(* Logix 5000 project; controller TFF vendor 1 type 14 code 107 rev 33.11; software revision 33.04; part 35 of 38 *)
(* tags used below, declared in another part *)
   Index : DINT;   // Index
   TIME : DINT[2];
   DigitalOutput : BOOL[256];   // Digital Output Array these bits are sent to output cards.
   FlowPath : FlowPath[64];   // Flow Path Array
   Options : Options;   // Options List
   PCV101_Control : PCV_Control;   // PCV101 Control UDT
   PCV201_Control : PCV_Control;   // PCV201 Control UDT
   PipeAnimation : PipeAnimation;   // HMI Pipe Animation Array
   PipeStatValueHMI : INT[224];   // Pipe Animation Value For HMI
   PTA001 : ALIAS FOR DigitalOutput[21];
   PTA101 : ALIAS FOR DigitalOutput[22];
   PTA201 : ALIAS FOR DigitalOutput[23];
   PTA401 : ALIAS FOR DigitalOutput[24];
   Rack_Murr_Node1_TFF20 : IO_Station;   // Status of Node 1 TFF20
   ThisSystem : SystemType;
   XV001 : ALIAS FOR Valve[0];
   XV002 : ALIAS FOR Valve[1];
   XV003 : ALIAS FOR Valve[2];
   XV004 : ALIAS FOR Valve[3];
   XV005 : ALIAS FOR Valve[4];
   XV006 : ALIAS FOR Valve[5];
   XV007 : ALIAS FOR Valve[6];
   XV101 : ALIAS FOR Valve[7];
   XV102 : ALIAS FOR Valve[8];
   XV201 : ALIAS FOR Valve[15];
   XV202 : ALIAS FOR Valve[16];
   XV401 : ALIAS FOR Valve[9];
   XV402 : ALIAS FOR Valve[10];
   XV403 : ALIAS FOR Valve[11];
   XV404 : ALIAS FOR Valve[12];
   XV405 : ALIAS FOR Valve[13];
   XV406 : ALIAS FOR Valve[14];
   XV701 : ALIAS FOR Valve[17];
   XV702 : ALIAS FOR Valve[18];
   XV703 : ALIAS FOR Valve[19];
   XV704 : ALIAS FOR Valve[20];
(* Process, continued *)

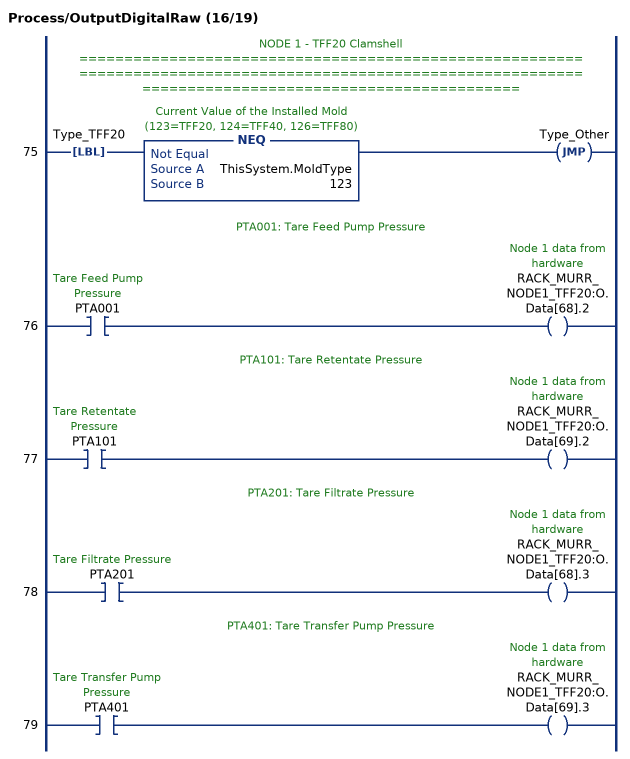
   // NODE 1 - TFF20 Clamshell
   // ==========================================================================================================================================================
   75: LBL(Type_TFF20)NEQ(ThisSystem.MoldType,123)JMP(Type_Other);
   // PTA001: Tare Feed Pump Pressure
   76: XIC(PTA001)OTE(RACK_MURR_NODE1_TFF20:O.Data[68].2);
   // PTA101: Tare Retentate Pressure
   77: XIC(PTA101)OTE(RACK_MURR_NODE1_TFF20:O.Data[69].2);
   // PTA201: Tare Filtrate Pressure
   78: XIC(PTA201)OTE(RACK_MURR_NODE1_TFF20:O.Data[68].3);
   // PTA401: Tare Transfer Pump Pressure
   79: XIC(PTA401)OTE(RACK_MURR_NODE1_TFF20:O.Data[69].3);
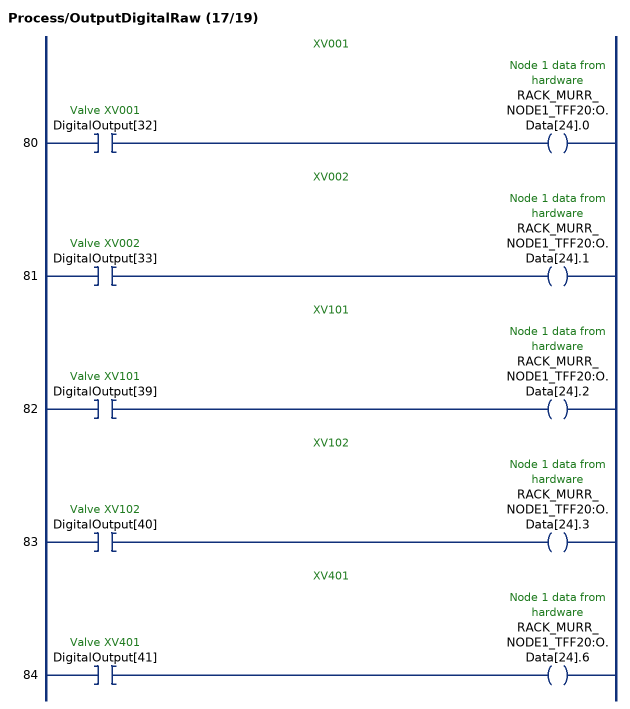
   // XV001
   80: XIC(DigitalOutput[32])OTE(RACK_MURR_NODE1_TFF20:O.Data[24].0);
   // XV002
   81: XIC(DigitalOutput[33])OTE(RACK_MURR_NODE1_TFF20:O.Data[24].1);
   // XV101
   82: XIC(DigitalOutput[39])OTE(RACK_MURR_NODE1_TFF20:O.Data[24].2);
   // XV102
   83: XIC(DigitalOutput[40])OTE(RACK_MURR_NODE1_TFF20:O.Data[24].3);
   // XV401
   84: XIC(DigitalOutput[41])OTE(RACK_MURR_NODE1_TFF20:O.Data[24].6);
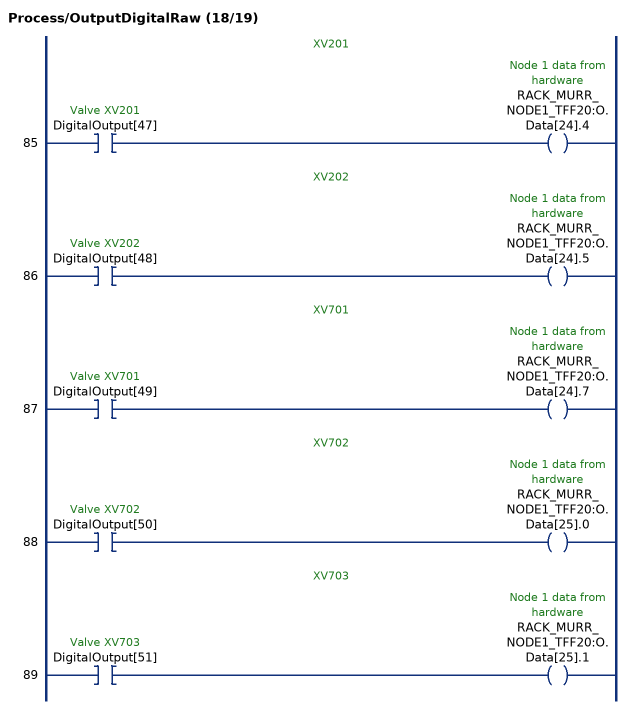
   // XV201
   85: XIC(DigitalOutput[47])OTE(RACK_MURR_NODE1_TFF20:O.Data[24].4);
   // XV202
   86: XIC(DigitalOutput[48])OTE(RACK_MURR_NODE1_TFF20:O.Data[24].5);
   // XV701
   87: XIC(DigitalOutput[49])OTE(RACK_MURR_NODE1_TFF20:O.Data[24].7);
   // XV702
   88: XIC(DigitalOutput[50])OTE(RACK_MURR_NODE1_TFF20:O.Data[25].0);
   // XV703
   89: XIC(DigitalOutput[51])OTE(RACK_MURR_NODE1_TFF20:O.Data[25].1);
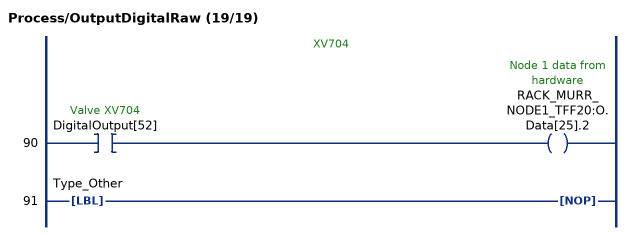
   // XV704
   90: XIC(DigitalOutput[52])OTE(RACK_MURR_NODE1_TFF20:O.Data[25].2);
   91: LBL(Type_Other)NOP();
END_ROUTINE

ROUTINE OutputProcessing   (* ladder *)
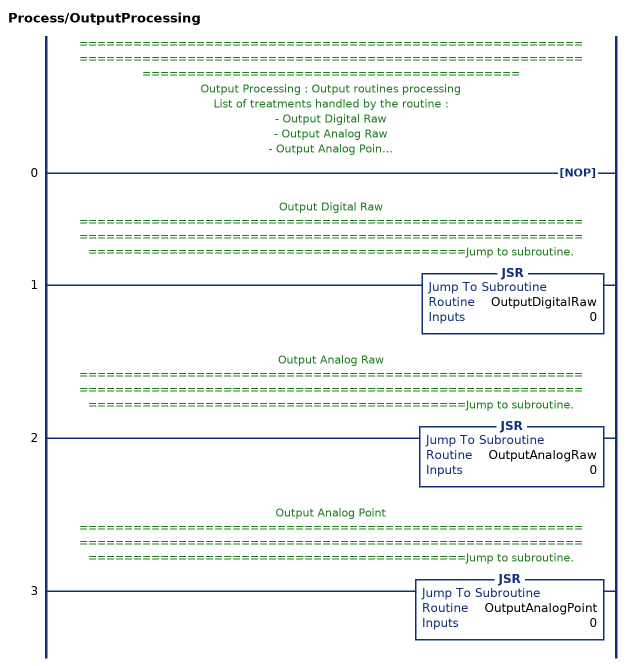
   // ==========================================================================================================================================================
   //                                                                                                                  Output Processing : Output routines processing
   //                                                     List of treatments handled by the routine :
   //                                                          - Output Digital Raw
   //                                                          - Output Analog Raw
   //                                                          - Output Analog Point
   //                                                     -----------------------------------------------------------------------------------------------------------------------------------------------------
   //                                                     History
   // 		2019-DEC-24 - Merck - Q. Spindler - Initial version for Candidate Release 1.00.00.00.a
   // ==========================================================================================================================================================
   0: NOP();
   // Output Digital Raw
   // ==========================================================================================================================================================Jump to subroutine.
   1: JSR(OutputDigitalRaw,0);
   // Output Analog Raw
   // ==========================================================================================================================================================Jump to subroutine.
   2: JSR(OutputAnalogRaw,0);
   // Output Analog Point
   // ==========================================================================================================================================================Jump to subroutine.
   3: JSR(OutputAnalogPoint,0);
END_ROUTINE

ROUTINE PipeAnimation   (* ladder *)
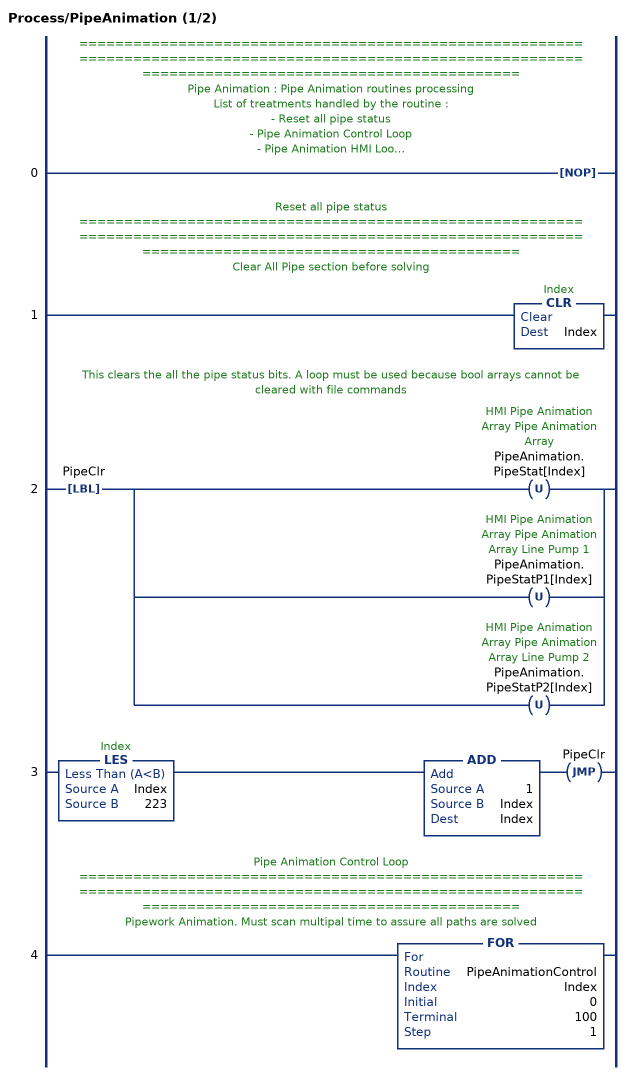
   // ==========================================================================================================================================================
   //                                                                                                               Pipe Animation : Pipe Animation routines processing
   //                                                     List of treatments handled by the routine :
   //                                                          - Reset all pipe status
   //                                                          - Pipe Animation Control Loop
   //                                                          - Pipe Animation HMI Loop
   //                                                     -----------------------------------------------------------------------------------------------------------------------------------------------------
   //                                                     History
   // 		2019-DEC-24 - Merck - Q. Spindler - Initial version for Candidate Release 1.00.00.00.a
   // ==========================================================================================================================================================
   0: NOP();
   // Reset all pipe status
   // ==========================================================================================================================================================
   // Clear All Pipe section before solving
   1: CLR(Index);
   // This clears the all the pipe status bits. A loop must be used because bool arrays cannot be cleared with file commands
   2: LBL(PipeClr)[OTU(PipeAnimation.PipeStat[Index]) ,OTU(PipeAnimation.PipeStatP1[Index]) ,OTU(PipeAnimation.PipeStatP2[Index]) ];
   3: LES(Index,223)ADD(1,Index,Index)JMP(PipeClr);
   // Pipe Animation Control Loop
   // ==========================================================================================================================================================
   // Pipework Animation. Must scan multipal time to assure all paths are solved
   4: FOR(PipeAnimationControl,Index,0,100,1);
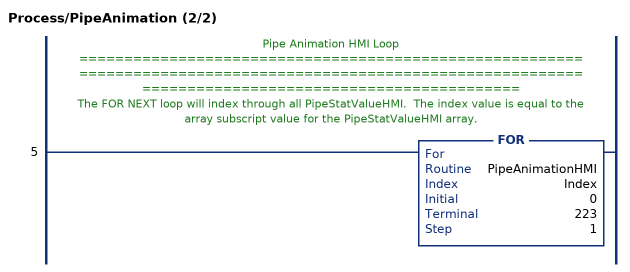
   // Pipe Animation HMI Loop
   // ==========================================================================================================================================================
   // The FOR NEXT loop will index through all PipeStatValueHMI.  The index value is equal to the array subscript value for the PipeStatValueHMI array.
   5: FOR(PipeAnimationHMI,Index,0,223,1);
END_ROUTINE

ROUTINE PipeAnimationControl   (* ladder *)
// Pipework Animation Routine
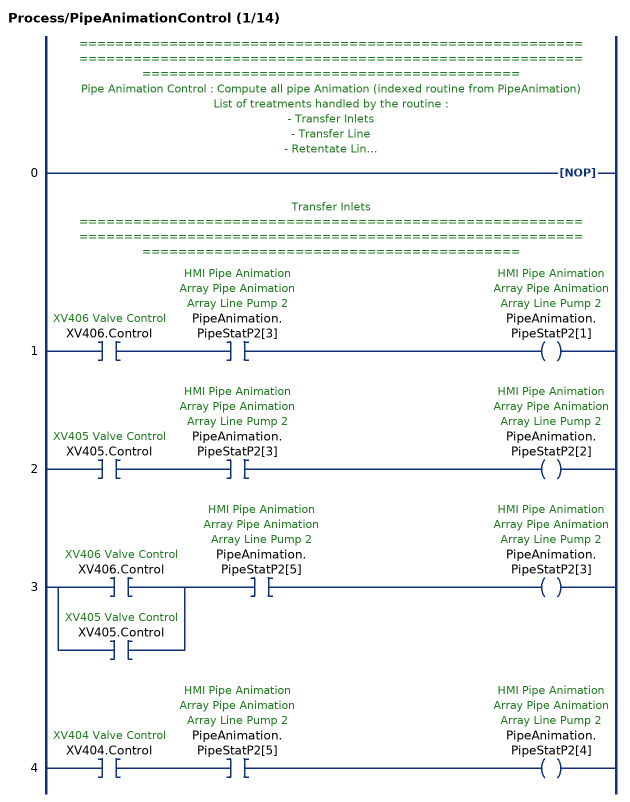
   // ==========================================================================================================================================================
   //                                                                                        Pipe Animation Control : Compute all pipe Animation (indexed routine from PipeAnimation)
   //                                                     List of treatments handled by the routine :
   //                                                          - Transfer Inlets
   //                                                          - Transfer Line
   //                                                          - Retentate Line
   //                                                           - Filtrate
   //                                                          - Feed Line
   //                                                           - Feed Inlets
   //                                                     -----------------------------------------------------------------------------------------------------------------------------------------------------
   //                                                     History
   // 		2019-DEC-24 - Merck - Q. Spindler - Initial version for Candidate Release 1.00.00.00.a
   // 		2020-JUN-19 - Merck - Q. Spindler - Modifications for Candidate Release 1.00.00.00.c
   //                                                                                             - Change State for Pipe ID 13, 14, 15, 16, 17, and 18 to prohibit Frontal filtration flowpath
   // ========================================================================================================================================================
   0: NOP();
   // Transfer Inlets
   // ==========================================================================================================================================================
   1: XIC(XV406.Control)XIC(PipeAnimation.PipeStatP2[3])OTE(PipeAnimation.PipeStatP2[1]);
   2: XIC(XV405.Control)XIC(PipeAnimation.PipeStatP2[3])OTE(PipeAnimation.PipeStatP2[2]);
   3: [XIC(XV406.Control) ,XIC(XV405.Control) ]XIC(PipeAnimation.PipeStatP2[5])OTE(PipeAnimation.PipeStatP2[3]);
   4: XIC(XV404.Control)XIC(PipeAnimation.PipeStatP2[5])OTE(PipeAnimation.PipeStatP2[4]);
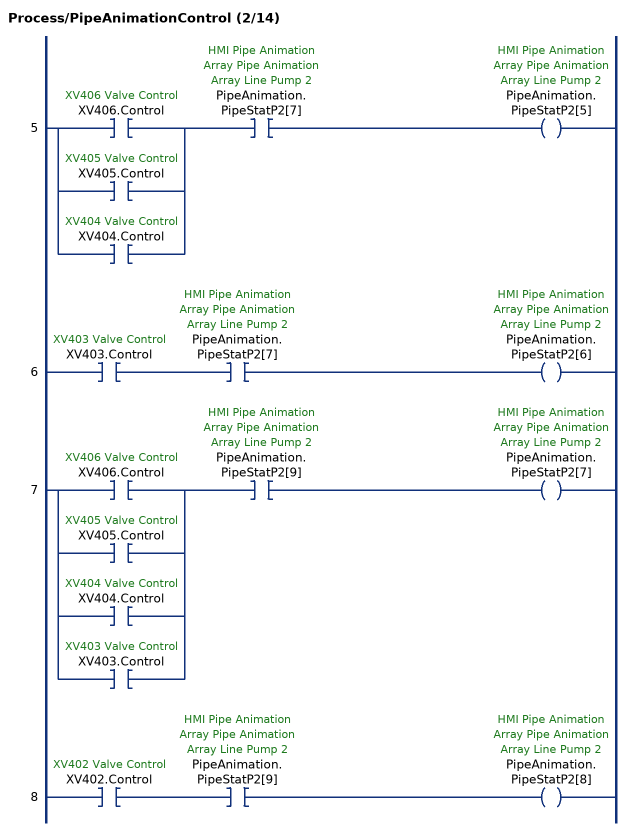
   5: [XIC(XV406.Control) ,XIC(XV405.Control) ,XIC(XV404.Control) ]XIC(PipeAnimation.PipeStatP2[7])OTE(PipeAnimation.PipeStatP2[5]);
   6: XIC(XV403.Control)XIC(PipeAnimation.PipeStatP2[7])OTE(PipeAnimation.PipeStatP2[6]);
   7: [XIC(XV406.Control) ,XIC(XV405.Control) ,XIC(XV404.Control) ,XIC(XV403.Control) ]XIC(PipeAnimation.PipeStatP2[9])OTE(PipeAnimation.PipeStatP2[7]);
   8: XIC(XV402.Control)XIC(PipeAnimation.PipeStatP2[9])OTE(PipeAnimation.PipeStatP2[8]);
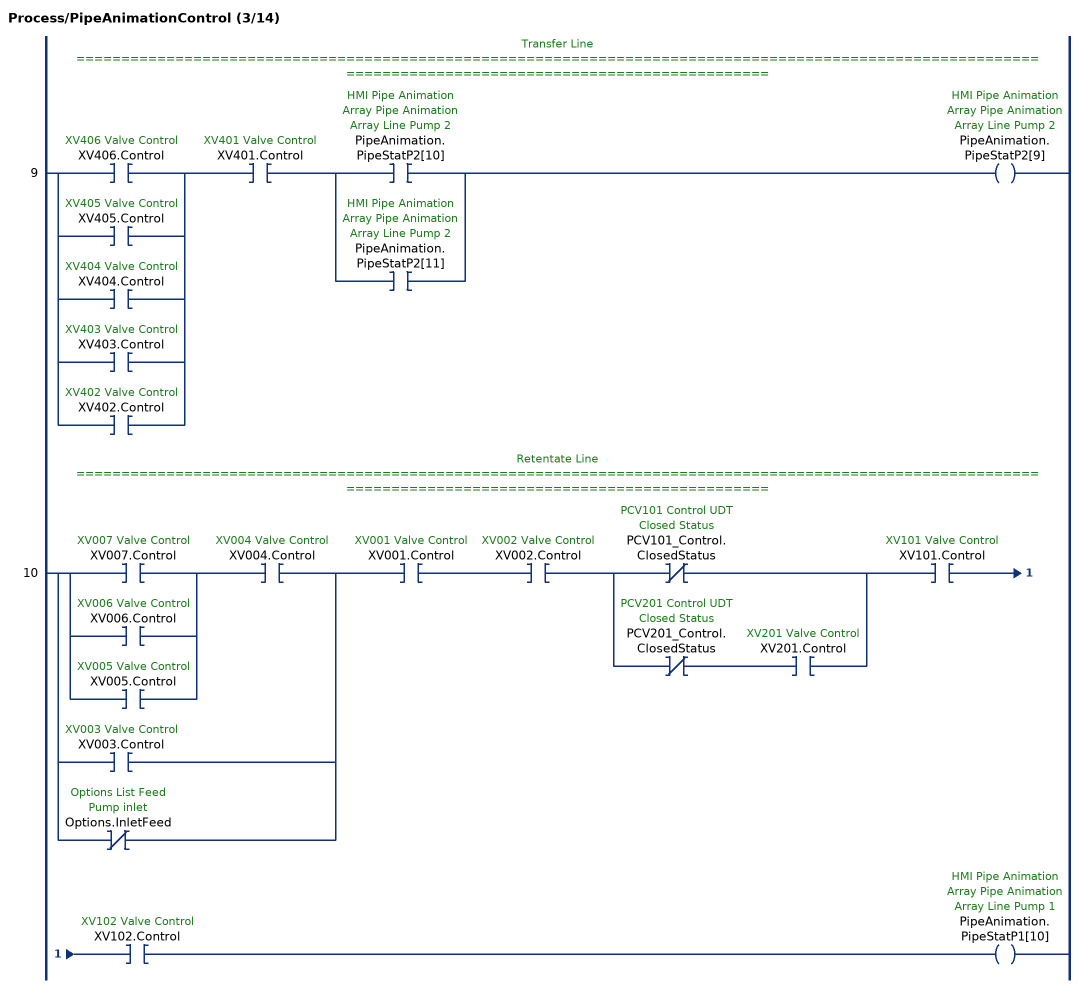
   // Transfer Line
   // ==========================================================================================================================================================
   9: [XIC(XV406.Control) ,XIC(XV405.Control) ,XIC(XV404.Control) ,XIC(XV403.Control) ,XIC(XV402.Control) ]XIC(XV401.Control)[XIC(PipeAnimation.PipeStatP2[10]) ,XIC(PipeAnimation.PipeStatP2[11]) ]OTE(PipeAnimation.PipeStatP2[9]);
   // Retentate Line
   // ==========================================================================================================================================================
   10: [[XIC(XV007.Control) ,XIC(XV006.Control) ,XIC(XV005.Control) ] XIC(XV004.Control) ,[XIC(XV003.Control) ,XIO(Options.InletFeed) ] ]XIC(XV001.Control)XIC(XV002.Control)[XIO(PCV101_Control.ClosedStatus) ,XIO(PCV201_Control.ClosedStatus) XIC(XV201.Control) ]XIC(XV101.Control)XIC(XV102.Control)OTE(PipeAnimation.PipeStatP1[10]);
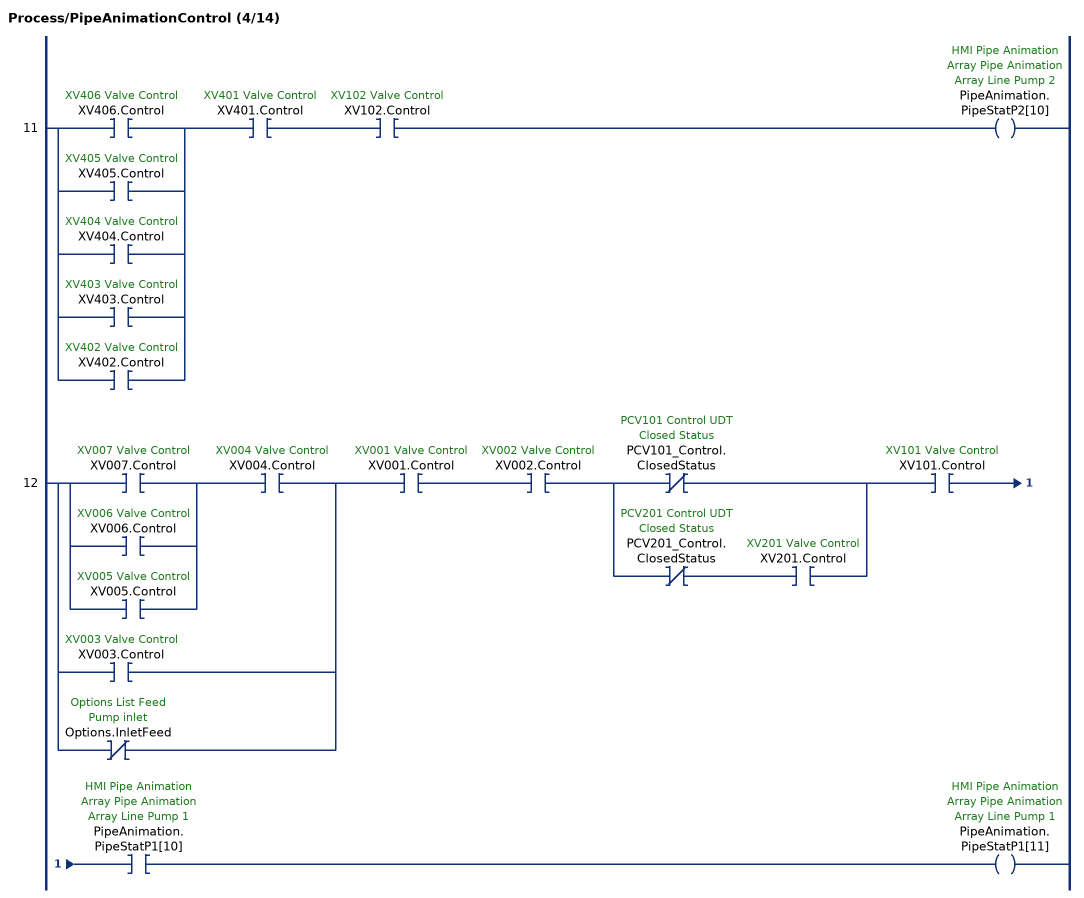
   11: [XIC(XV406.Control) ,XIC(XV405.Control) ,XIC(XV404.Control) ,XIC(XV403.Control) ,XIC(XV402.Control) ]XIC(XV401.Control)XIC(XV102.Control)OTE(PipeAnimation.PipeStatP2[10]);
   12: [[XIC(XV007.Control) ,XIC(XV006.Control) ,XIC(XV005.Control) ] XIC(XV004.Control) ,[XIC(XV003.Control) ,XIO(Options.InletFeed) ] ]XIC(XV001.Control)XIC(XV002.Control)[XIO(PCV101_Control.ClosedStatus) ,XIO(PCV201_Control.ClosedStatus) XIC(XV201.Control) ]XIC(XV101.Control)XIC(PipeAnimation.PipeStatP1[10])OTE(PipeAnimation.PipeStatP1[11]);
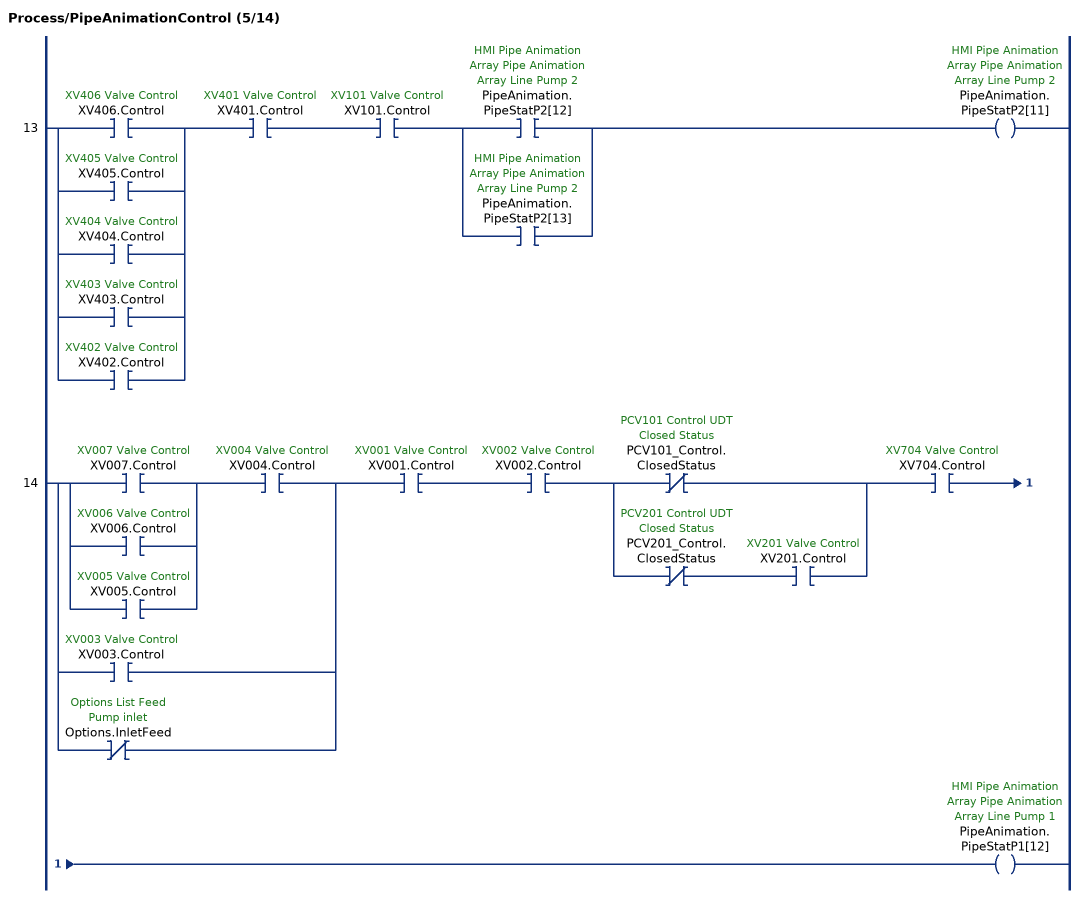
   13: [XIC(XV406.Control) ,XIC(XV405.Control) ,XIC(XV404.Control) ,XIC(XV403.Control) ,XIC(XV402.Control) ]XIC(XV401.Control)XIC(XV101.Control)[XIC(PipeAnimation.PipeStatP2[12]) ,XIC(PipeAnimation.PipeStatP2[13]) ]OTE(PipeAnimation.PipeStatP2[11]);
   14: [[XIC(XV007.Control) ,XIC(XV006.Control) ,XIC(XV005.Control) ] XIC(XV004.Control) ,[XIC(XV003.Control) ,XIO(Options.InletFeed) ] ]XIC(XV001.Control)XIC(XV002.Control)[XIO(PCV101_Control.ClosedStatus) ,XIO(PCV201_Control.ClosedStatus) XIC(XV201.Control) ]XIC(XV704.Control)OTE(PipeAnimation.PipeStatP1[12]);
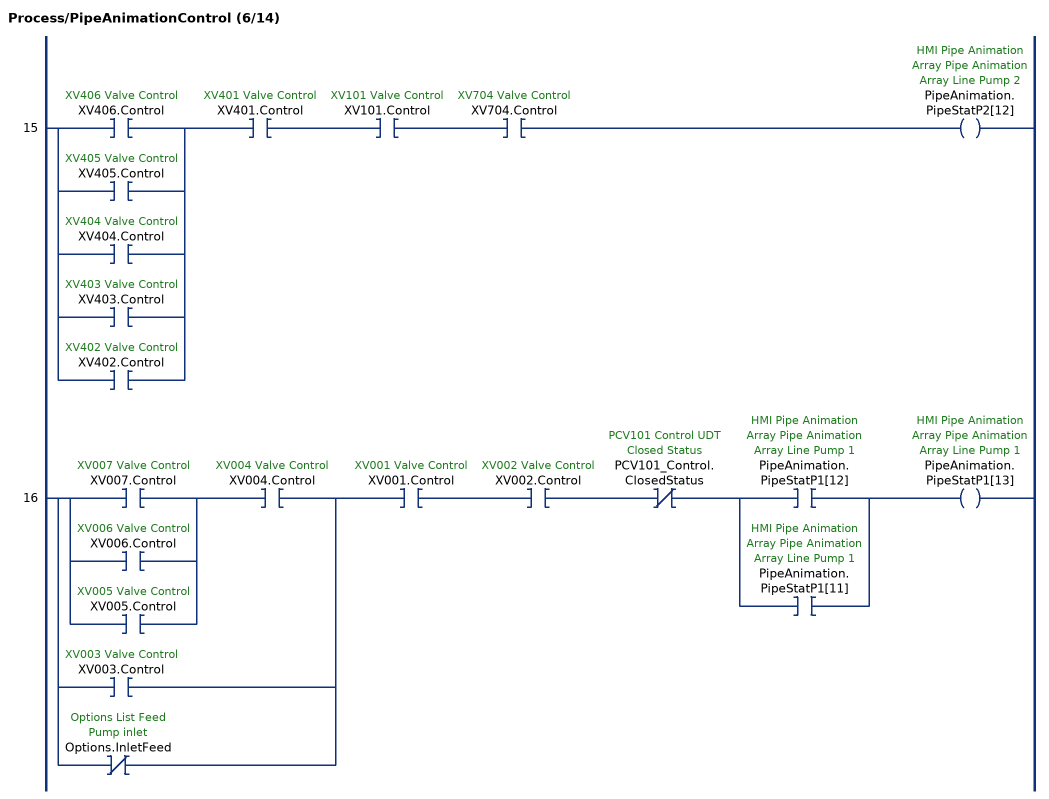
   15: [XIC(XV406.Control) ,XIC(XV405.Control) ,XIC(XV404.Control) ,XIC(XV403.Control) ,XIC(XV402.Control) ]XIC(XV401.Control)XIC(XV101.Control)XIC(XV704.Control)OTE(PipeAnimation.PipeStatP2[12]);
   16: [[XIC(XV007.Control) ,XIC(XV006.Control) ,XIC(XV005.Control) ] XIC(XV004.Control) ,[XIC(XV003.Control) ,XIO(Options.InletFeed) ] ]XIC(XV001.Control)XIC(XV002.Control)XIO(PCV101_Control.ClosedStatus)[XIC(PipeAnimation.PipeStatP1[12]) ,XIC(PipeAnimation.PipeStatP1[11]) ]OTE(PipeAnimation.PipeStatP1[13]);
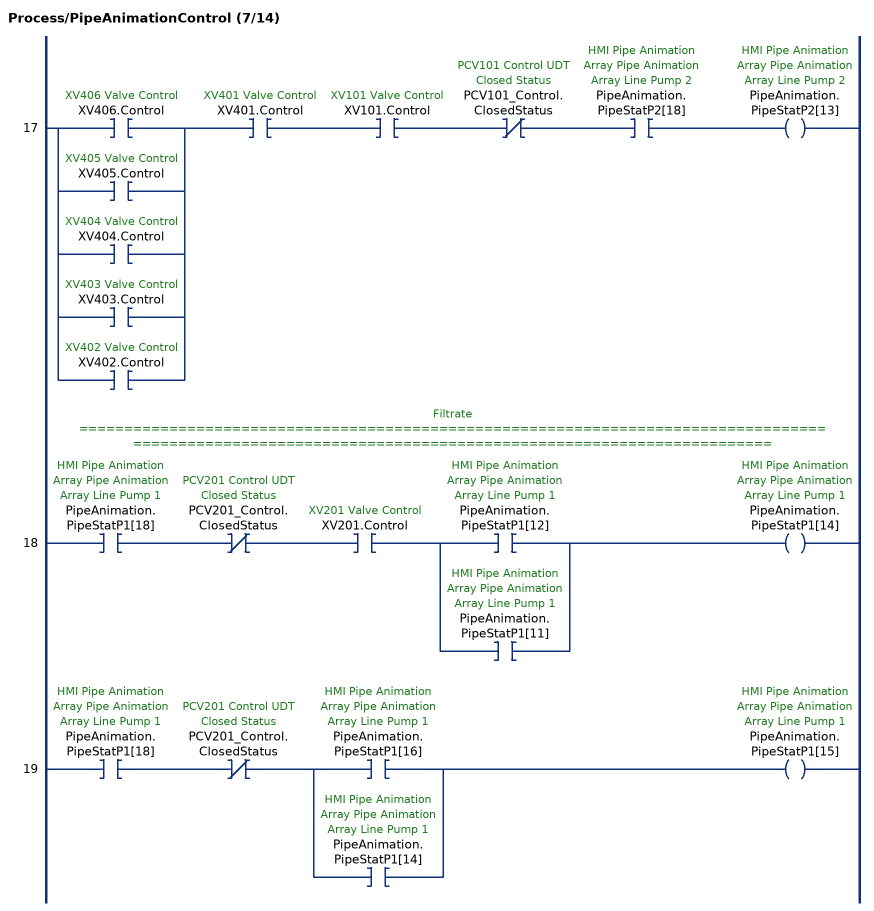
   17: [XIC(XV406.Control) ,XIC(XV405.Control) ,XIC(XV404.Control) ,XIC(XV403.Control) ,XIC(XV402.Control) ]XIC(XV401.Control)XIC(XV101.Control)XIO(PCV101_Control.ClosedStatus)XIC(PipeAnimation.PipeStatP2[18])OTE(PipeAnimation.PipeStatP2[13]);
   // Filtrate
   // ==========================================================================================================================================================
   18: XIC(PipeAnimation.PipeStatP1[18])XIO(PCV201_Control.ClosedStatus)XIC(XV201.Control)[XIC(PipeAnimation.PipeStatP1[12]) ,XIC(PipeAnimation.PipeStatP1[11]) ]OTE(PipeAnimation.PipeStatP1[14]);
   19: XIC(PipeAnimation.PipeStatP1[18])XIO(PCV201_Control.ClosedStatus)[XIC(PipeAnimation.PipeStatP1[16]) ,XIC(PipeAnimation.PipeStatP1[14]) ]OTE(PipeAnimation.PipeStatP1[15]);
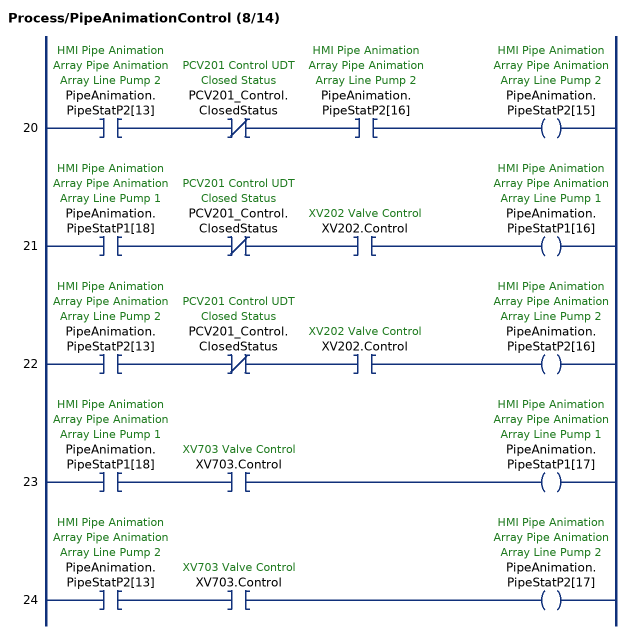
   20: XIC(PipeAnimation.PipeStatP2[13])XIO(PCV201_Control.ClosedStatus)XIC(PipeAnimation.PipeStatP2[16])OTE(PipeAnimation.PipeStatP2[15]);
   21: XIC(PipeAnimation.PipeStatP1[18])XIO(PCV201_Control.ClosedStatus)XIC(XV202.Control)OTE(PipeAnimation.PipeStatP1[16]);
   22: XIC(PipeAnimation.PipeStatP2[13])XIO(PCV201_Control.ClosedStatus)XIC(XV202.Control)OTE(PipeAnimation.PipeStatP2[16]);
   23: XIC(PipeAnimation.PipeStatP1[18])XIC(XV703.Control)OTE(PipeAnimation.PipeStatP1[17]);
   24: XIC(PipeAnimation.PipeStatP2[13])XIC(XV703.Control)OTE(PipeAnimation.PipeStatP2[17]);
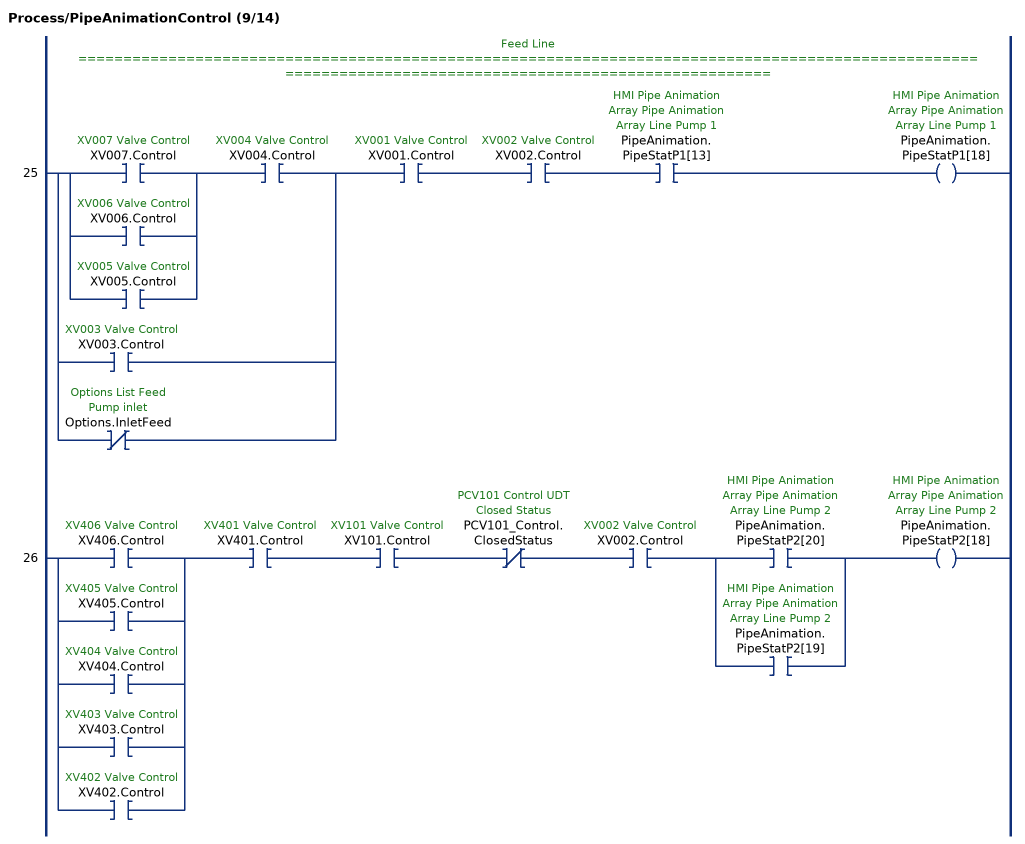
   // Feed Line
   // ==========================================================================================================================================================
   25: [[XIC(XV007.Control) ,XIC(XV006.Control) ,XIC(XV005.Control) ] XIC(XV004.Control) ,[XIC(XV003.Control) ,XIO(Options.InletFeed) ] ]XIC(XV001.Control)XIC(XV002.Control)XIC(PipeAnimation.PipeStatP1[13])OTE(PipeAnimation.PipeStatP1[18]);
   26: [XIC(XV406.Control) ,XIC(XV405.Control) ,XIC(XV404.Control) ,XIC(XV403.Control) ,XIC(XV402.Control) ]XIC(XV401.Control)XIC(XV101.Control)XIO(PCV101_Control.ClosedStatus)XIC(XV002.Control)[XIC(PipeAnimation.PipeStatP2[20]) ,XIC(PipeAnimation.PipeStatP2[19]) ]OTE(PipeAnimation.PipeStatP2[18]);
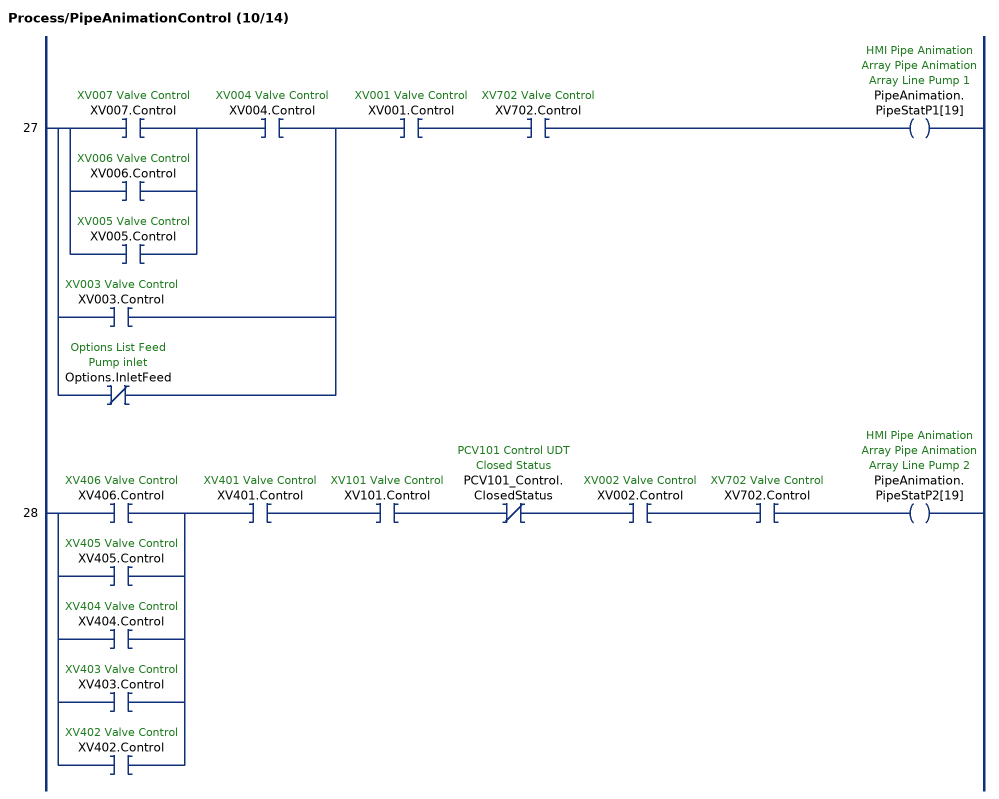
   27: [[XIC(XV007.Control) ,XIC(XV006.Control) ,XIC(XV005.Control) ] XIC(XV004.Control) ,[XIC(XV003.Control) ,XIO(Options.InletFeed) ] ]XIC(XV001.Control)XIC(XV702.Control)OTE(PipeAnimation.PipeStatP1[19]);
   28: [XIC(XV406.Control) ,XIC(XV405.Control) ,XIC(XV404.Control) ,XIC(XV403.Control) ,XIC(XV402.Control) ]XIC(XV401.Control)XIC(XV101.Control)XIO(PCV101_Control.ClosedStatus)XIC(XV002.Control)XIC(XV702.Control)OTE(PipeAnimation.PipeStatP2[19]);
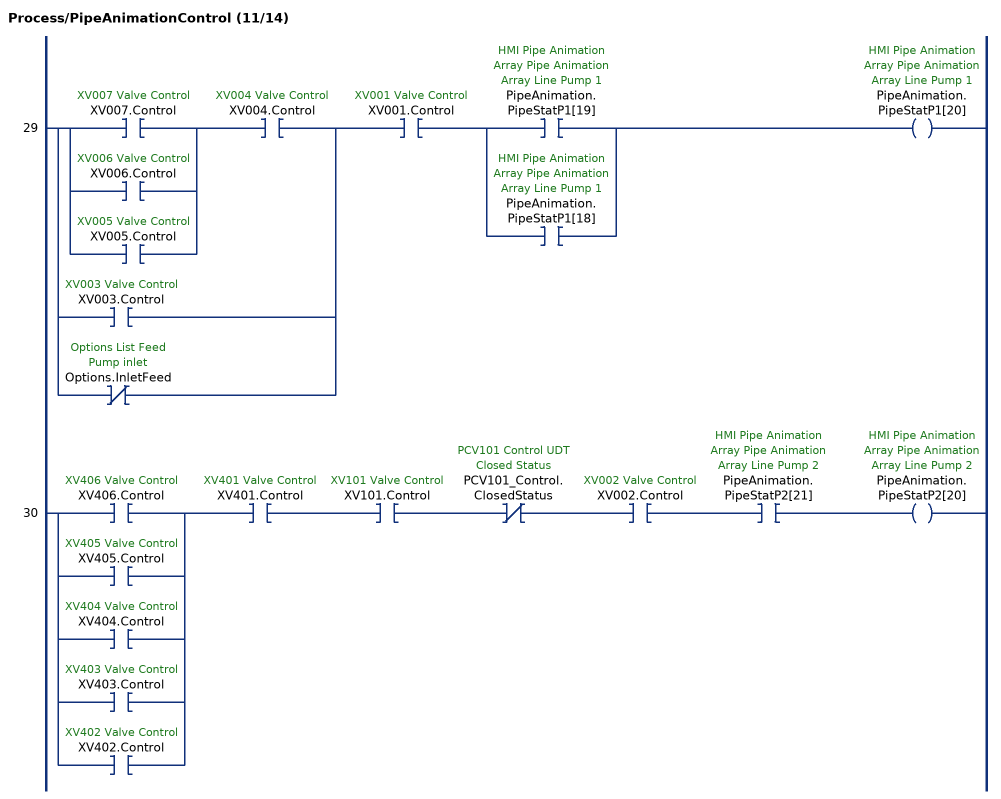
   29: [[XIC(XV007.Control) ,XIC(XV006.Control) ,XIC(XV005.Control) ] XIC(XV004.Control) ,[XIC(XV003.Control) ,XIO(Options.InletFeed) ] ]XIC(XV001.Control)[XIC(PipeAnimation.PipeStatP1[19]) ,XIC(PipeAnimation.PipeStatP1[18]) ]OTE(PipeAnimation.PipeStatP1[20]);
   30: [XIC(XV406.Control) ,XIC(XV405.Control) ,XIC(XV404.Control) ,XIC(XV403.Control) ,XIC(XV402.Control) ]XIC(XV401.Control)XIC(XV101.Control)XIO(PCV101_Control.ClosedStatus)XIC(XV002.Control)XIC(PipeAnimation.PipeStatP2[21])OTE(PipeAnimation.PipeStatP2[20]);
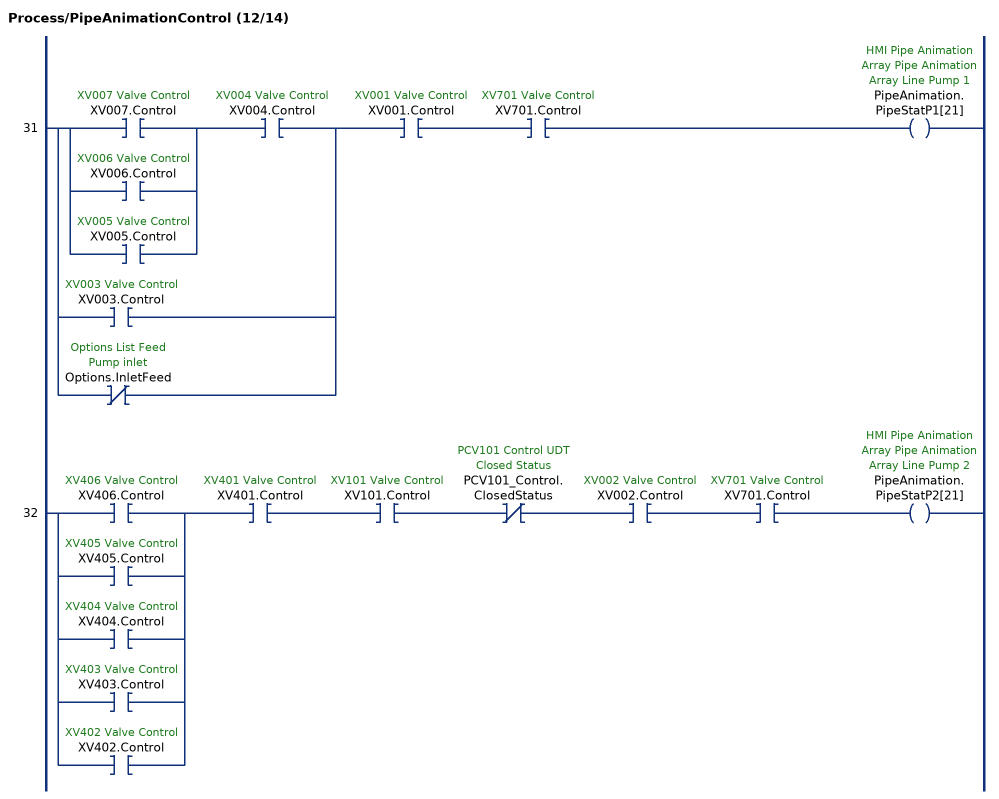
   31: [[XIC(XV007.Control) ,XIC(XV006.Control) ,XIC(XV005.Control) ] XIC(XV004.Control) ,[XIC(XV003.Control) ,XIO(Options.InletFeed) ] ]XIC(XV001.Control)XIC(XV701.Control)OTE(PipeAnimation.PipeStatP1[21]);
   32: [XIC(XV406.Control) ,XIC(XV405.Control) ,XIC(XV404.Control) ,XIC(XV403.Control) ,XIC(XV402.Control) ]XIC(XV401.Control)XIC(XV101.Control)XIO(PCV101_Control.ClosedStatus)XIC(XV002.Control)XIC(XV701.Control)OTE(PipeAnimation.PipeStatP2[21]);
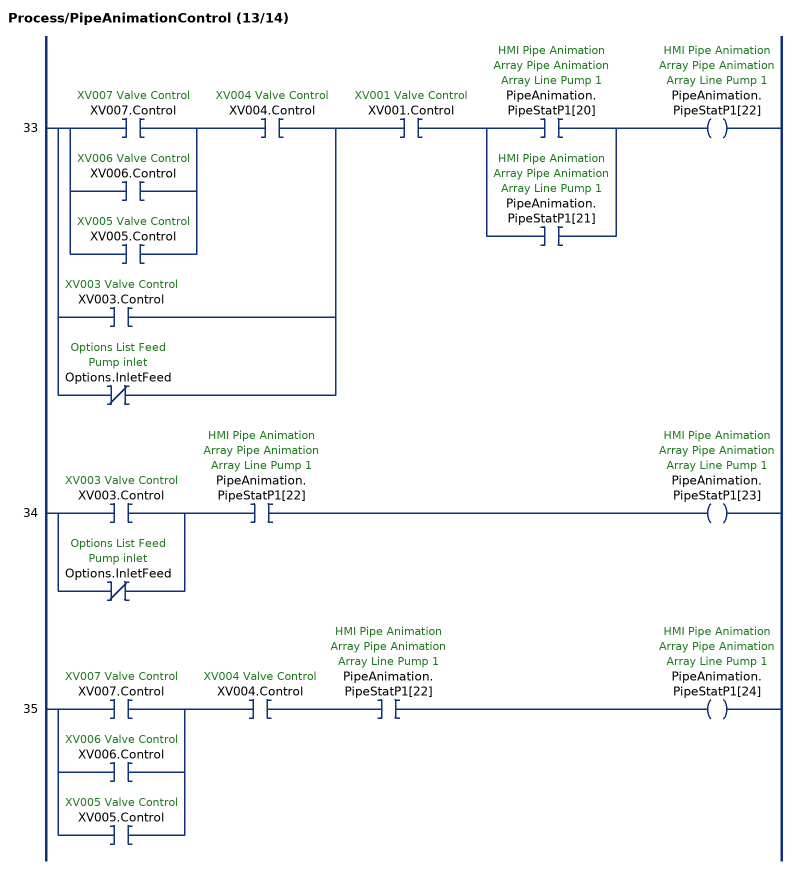
   33: [[XIC(XV007.Control) ,XIC(XV006.Control) ,XIC(XV005.Control) ] XIC(XV004.Control) ,[XIC(XV003.Control) ,XIO(Options.InletFeed) ] ]XIC(XV001.Control)[XIC(PipeAnimation.PipeStatP1[20]) ,XIC(PipeAnimation.PipeStatP1[21]) ]OTE(PipeAnimation.PipeStatP1[22]);
   34: [XIC(XV003.Control) ,XIO(Options.InletFeed) ]XIC(PipeAnimation.PipeStatP1[22])OTE(PipeAnimation.PipeStatP1[23]);
   35: [XIC(XV007.Control) ,XIC(XV006.Control) ,XIC(XV005.Control) ]XIC(XV004.Control)XIC(PipeAnimation.PipeStatP1[22])OTE(PipeAnimation.PipeStatP1[24]);
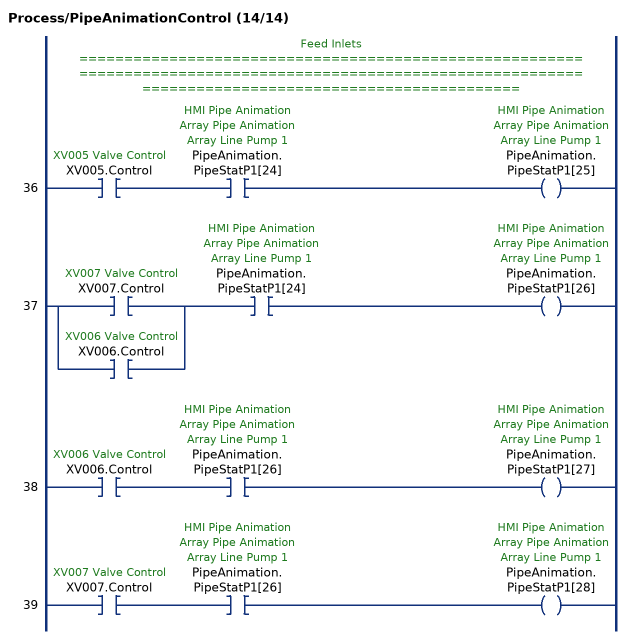
   // Feed Inlets
   // ==========================================================================================================================================================
   36: XIC(XV005.Control)XIC(PipeAnimation.PipeStatP1[24])OTE(PipeAnimation.PipeStatP1[25]);
   37: [XIC(XV007.Control) ,XIC(XV006.Control) ]XIC(PipeAnimation.PipeStatP1[24])OTE(PipeAnimation.PipeStatP1[26]);
   38: XIC(XV006.Control)XIC(PipeAnimation.PipeStatP1[26])OTE(PipeAnimation.PipeStatP1[27]);
   39: XIC(XV007.Control)XIC(PipeAnimation.PipeStatP1[26])OTE(PipeAnimation.PipeStatP1[28]);
END_ROUTINE
